// Tests for HalfBROT.FB_FocusManualHome, the decision and the end detection of a manual focus re-home, calibrated or not (HalfBROT 0.11.0, #138).
// The wiring in FB_FocusControl and the NC behaviour are not testable here (the mock skips the body): on-site test.
FUNCTION_BLOCK FB_FocusManualHome_Tests EXTENDS TcUnit.FB_TestSuite
VAR
END_VAR

Accepted_When_Calibrated_Idle_Automatic();
Rejected_In_Manual_Mode();
Rejected_With_Manual_Unlock();
Rejected_With_Axis_Error();
Accepted_When_Not_Calibrated();
Uncalibrated_Rejected_In_Manual_Mode();
Uncalibrated_Rejected_While_Homing();
Uncalibrated_Rejected_With_Error();
Uncalibrated_Rejected_With_Manual_Unlock();
Uncalibrated_Rejected_While_Moving();
NotAutomatic_Before_Homing();
No_Second_Request_While_Running_Uncalibrated();
Calibrated_Request_Restores_Target();
Uncalibrated_Done_No_Restore();
Uncalibrated_Abort_Blocks_AutoHome();
Uncalibrated_Abort_Before_Start();
Rejected_While_Homing();
Rejected_While_Moving();
No_Second_Request_While_Running();
Done_After_Active_And_Calibrated();
Done_When_Calibrated_Stays_True();
Done_When_Calibrated_Drops_And_Returns();
Abort_By_Stop_Pulse();
Abort_By_Error();
Abort_Before_Start();
Abort_Uncalibrated_Blocks_AutoHome();
Abort_Calibrated_No_Block();
Request_Clears_Block();
ClearBlock();
Aborted_Rehome_Then_Rehome_Restores_The_First_Target();
ClearBlock_Drops_The_Kept_Target();
Calibrated_Abort_Drops_The_Pending_Target();

// The plain case: accepted, running, the target is kept for the end.
METHOD PRIVATE Accepted_When_Calibrated_Idle_Automatic
VAR
	fb	: HalfBROT.FB_FocusManualHome;
	eRes	: HalfBROT.E_FocusManualHome;
END_VAR
TEST('Accepted_When_Calibrated_Idle_Automatic');
eRes := fb.Request(bAutomatic := TRUE, bManualUnlock := FALSE, bError := FALSE, bCalibrated := TRUE, bHoming := FALSE, bMoving := FALSE, fTarget := 36.0);
AssertTrue(Condition := eRes = HalfBROT.E_FocusManualHome.Accepted, Message := 'accepted');
AssertTrue(Condition := fb.bRunning, Message := 'running');
AssertFalse(Condition := fb.bBlockAutoHome, Message := 'no block');
AssertEquals_LREAL(Expected := 36.0, Actual := fb.fRestoreTarget, Delta := 1.0E-9, Message := 'target kept');
AssertTrue(Condition := fb.bRestoreTarget, Message := 'restore the target');
TEST_FINISHED();
END_METHOD

// Manual/pendant mode: the pendant drives the enable and jogs.
METHOD PRIVATE Rejected_In_Manual_Mode
VAR
	fb	: HalfBROT.FB_FocusManualHome;
	eRes	: HalfBROT.E_FocusManualHome;
END_VAR
TEST('Rejected_In_Manual_Mode');
eRes := fb.Request(bAutomatic := FALSE, bManualUnlock := FALSE, bError := FALSE, bCalibrated := TRUE, bHoming := FALSE, bMoving := FALSE, fTarget := 36.0);
AssertTrue(Condition := eRes = HalfBROT.E_FocusManualHome.NotAutomatic, Message := 'manual mode');
AssertFalse(Condition := fb.bRunning, Message := 'nothing started');
TEST_FINISHED();
END_METHOD

METHOD PRIVATE Rejected_With_Manual_Unlock
VAR
	fb	: HalfBROT.FB_FocusManualHome;
	eRes	: HalfBROT.E_FocusManualHome;
END_VAR
TEST('Rejected_With_Manual_Unlock');
eRes := fb.Request(bAutomatic := TRUE, bManualUnlock := TRUE, bError := FALSE, bCalibrated := TRUE, bHoming := FALSE, bMoving := FALSE, fTarget := 36.0);
AssertTrue(Condition := eRes = HalfBROT.E_FocusManualHome.ManualUnlock, Message := 'manual unlock');
AssertFalse(Condition := fb.bRunning, Message := 'nothing started');
TEST_FINISHED();
END_METHOD

METHOD PRIVATE Rejected_With_Axis_Error
VAR
	fb	: HalfBROT.FB_FocusManualHome;
	eRes	: HalfBROT.E_FocusManualHome;
END_VAR
TEST('Rejected_With_Axis_Error');
eRes := fb.Request(bAutomatic := TRUE, bManualUnlock := FALSE, bError := TRUE, bCalibrated := TRUE, bHoming := FALSE, bMoving := FALSE, fTarget := 36.0);
AssertTrue(Condition := eRes = HalfBROT.E_FocusManualHome.AxisError, Message := 'axis error');
AssertFalse(Condition := fb.bRunning, Message := 'nothing started');
TEST_FINISHED();
END_METHOD

// A homing is requested, pending or active (the caller passes bHomeAxis OR HomeActive OR HomePending).
METHOD PRIVATE Rejected_While_Homing
VAR
	fb	: HalfBROT.FB_FocusManualHome;
	eRes	: HalfBROT.E_FocusManualHome;
END_VAR
TEST('Rejected_While_Homing');
eRes := fb.Request(bAutomatic := TRUE, bManualUnlock := FALSE, bError := FALSE, bCalibrated := TRUE, bHoming := TRUE, bMoving := FALSE, fTarget := 36.0);
AssertTrue(Condition := eRes = HalfBROT.E_FocusManualHome.Homing, Message := 'homing');
AssertFalse(Condition := fb.bRunning, Message := 'nothing started');
TEST_FINISHED();
END_METHOD

METHOD PRIVATE Rejected_While_Moving
VAR
	fb	: HalfBROT.FB_FocusManualHome;
	eRes	: HalfBROT.E_FocusManualHome;
END_VAR
TEST('Rejected_While_Moving');
eRes := fb.Request(bAutomatic := TRUE, bManualUnlock := FALSE, bError := FALSE, bCalibrated := TRUE, bHoming := FALSE, bMoving := TRUE, fTarget := 36.0);
AssertTrue(Condition := eRes = HalfBROT.E_FocusManualHome.Moving, Message := 'moving');
AssertFalse(Condition := fb.bRunning, Message := 'nothing started');
TEST_FINISHED();
END_METHOD

METHOD PRIVATE No_Second_Request_While_Running
VAR
	fb	: HalfBROT.FB_FocusManualHome;
	eRes	: HalfBROT.E_FocusManualHome;
END_VAR
TEST('No_Second_Request_While_Running');
eRes := fb.Request(bAutomatic := TRUE, bManualUnlock := FALSE, bError := FALSE, bCalibrated := TRUE, bHoming := FALSE, bMoving := FALSE, fTarget := 36.0);
eRes := fb.Request(bAutomatic := TRUE, bManualUnlock := FALSE, bError := FALSE, bCalibrated := TRUE, bHoming := FALSE, bMoving := FALSE, fTarget := 50.0);
AssertTrue(Condition := eRes = HalfBROT.E_FocusManualHome.Homing, Message := 'second request');
AssertEquals_LREAL(Expected := 36.0, Actual := fb.fRestoreTarget, Delta := 1.0E-9, Message := 'first target kept');
TEST_FINISHED();
END_METHOD

// Pending, active, then calibrated and idle: done for one cycle, restore target available.
METHOD PRIVATE Done_After_Active_And_Calibrated
VAR
	fb	: HalfBROT.FB_FocusManualHome;
	eRes	: HalfBROT.E_FocusManualHome;
END_VAR
TEST('Done_After_Active_And_Calibrated');
eRes := fb.Request(bAutomatic := TRUE, bManualUnlock := FALSE, bError := FALSE, bCalibrated := TRUE, bHoming := FALSE, bMoving := FALSE, fTarget := 36.0);
fb(bHomeActive := FALSE, bHomePending := TRUE, bCalibrated := TRUE, bAbortPulse := FALSE);
AssertTrue(Condition := fb.bRunning, Message := 'running while pending');
fb(bHomeActive := TRUE, bHomePending := FALSE, bCalibrated := TRUE, bAbortPulse := FALSE);
AssertTrue(Condition := fb.bRunning, Message := 'running while active');
AssertFalse(Condition := fb.bDone, Message := 'not done yet');
fb(bHomeActive := FALSE, bHomePending := FALSE, bCalibrated := TRUE, bAbortPulse := FALSE);
AssertTrue(Condition := fb.bDone, Message := 'done');
AssertFalse(Condition := fb.bRunning, Message := 'ended');
AssertFalse(Condition := fb.bAborted, Message := 'not aborted');
AssertFalse(Condition := fb.bBlockAutoHome, Message := 'no block');
fb(bHomeActive := FALSE, bHomePending := FALSE, bCalibrated := TRUE, bAbortPulse := FALSE);
AssertFalse(Condition := fb.bDone, Message := 'done is one cycle');
TEST_FINISHED();
END_METHOD

// The NC keeps Homed during the homing.
METHOD PRIVATE Done_When_Calibrated_Stays_True
VAR
	fb	: HalfBROT.FB_FocusManualHome;
	eRes	: HalfBROT.E_FocusManualHome;
END_VAR
TEST('Done_When_Calibrated_Stays_True');
eRes := fb.Request(bAutomatic := TRUE, bManualUnlock := FALSE, bError := FALSE, bCalibrated := TRUE, bHoming := FALSE, bMoving := FALSE, fTarget := 36.0);
fb(bHomeActive := TRUE, bHomePending := FALSE, bCalibrated := TRUE, bAbortPulse := FALSE);
fb(bHomeActive := TRUE, bHomePending := FALSE, bCalibrated := TRUE, bAbortPulse := FALSE);
fb(bHomeActive := FALSE, bHomePending := FALSE, bCalibrated := TRUE, bAbortPulse := FALSE);
AssertTrue(Condition := fb.bDone, Message := 'done');
TEST_FINISHED();
END_METHOD

// The NC drops Homed at the start of the homing.
METHOD PRIVATE Done_When_Calibrated_Drops_And_Returns
VAR
	fb	: HalfBROT.FB_FocusManualHome;
	eRes	: HalfBROT.E_FocusManualHome;
END_VAR
TEST('Done_When_Calibrated_Drops_And_Returns');
eRes := fb.Request(bAutomatic := TRUE, bManualUnlock := FALSE, bError := FALSE, bCalibrated := TRUE, bHoming := FALSE, bMoving := FALSE, fTarget := 36.0);
fb(bHomeActive := FALSE, bHomePending := TRUE, bCalibrated := TRUE, bAbortPulse := FALSE);
fb(bHomeActive := TRUE, bHomePending := FALSE, bCalibrated := FALSE, bAbortPulse := FALSE);
fb(bHomeActive := TRUE, bHomePending := FALSE, bCalibrated := FALSE, bAbortPulse := FALSE);
fb(bHomeActive := FALSE, bHomePending := FALSE, bCalibrated := TRUE, bAbortPulse := FALSE);
AssertTrue(Condition := fb.bDone, Message := 'done');
AssertFalse(Condition := fb.bBlockAutoHome, Message := 'no block');
TEST_FINISHED();
END_METHOD

// A stop aborts the homing; the axis keeps its old calibration.
METHOD PRIVATE Abort_By_Stop_Pulse
VAR
	fb	: HalfBROT.FB_FocusManualHome;
	eRes	: HalfBROT.E_FocusManualHome;
END_VAR
TEST('Abort_By_Stop_Pulse');
eRes := fb.Request(bAutomatic := TRUE, bManualUnlock := FALSE, bError := FALSE, bCalibrated := TRUE, bHoming := FALSE, bMoving := FALSE, fTarget := 36.0);
fb(bHomeActive := TRUE, bHomePending := FALSE, bCalibrated := TRUE, bAbortPulse := FALSE);
fb(bHomeActive := TRUE, bHomePending := FALSE, bCalibrated := TRUE, bAbortPulse := TRUE);
fb(bHomeActive := FALSE, bHomePending := FALSE, bCalibrated := TRUE, bAbortPulse := FALSE);
AssertTrue(Condition := fb.bAborted, Message := 'aborted');
AssertFalse(Condition := fb.bDone, Message := 'not done');
AssertFalse(Condition := fb.bRunning, Message := 'ended');
AssertFalse(Condition := fb.bBlockAutoHome, Message := 'calibrated: no block');
TEST_FINISHED();
END_METHOD

// An axis error ends the homing uncalibrated.
METHOD PRIVATE Abort_By_Error
VAR
	fb	: HalfBROT.FB_FocusManualHome;
	eRes	: HalfBROT.E_FocusManualHome;
END_VAR
TEST('Abort_By_Error');
eRes := fb.Request(bAutomatic := TRUE, bManualUnlock := FALSE, bError := FALSE, bCalibrated := TRUE, bHoming := FALSE, bMoving := FALSE, fTarget := 36.0);
fb(bHomeActive := TRUE, bHomePending := FALSE, bCalibrated := TRUE, bAbortPulse := FALSE);
fb(bHomeActive := TRUE, bHomePending := FALSE, bCalibrated := FALSE, bAbortPulse := TRUE);
fb(bHomeActive := FALSE, bHomePending := FALSE, bCalibrated := FALSE, bAbortPulse := FALSE);
AssertTrue(Condition := fb.bAborted, Message := 'aborted');
AssertFalse(Condition := fb.bDone, Message := 'not done');
AssertTrue(Condition := fb.bBlockAutoHome, Message := 'uncalibrated: block');
TEST_FINISHED();
END_METHOD

// Stop() cancels a Home() that still waits for the drive: HomeActive is never seen.
METHOD PRIVATE Abort_Before_Start
VAR
	fb	: HalfBROT.FB_FocusManualHome;
	eRes	: HalfBROT.E_FocusManualHome;
END_VAR
TEST('Abort_Before_Start');
eRes := fb.Request(bAutomatic := TRUE, bManualUnlock := FALSE, bError := FALSE, bCalibrated := TRUE, bHoming := FALSE, bMoving := FALSE, fTarget := 36.0);
fb(bHomeActive := FALSE, bHomePending := TRUE, bCalibrated := TRUE, bAbortPulse := FALSE);
fb(bHomeActive := FALSE, bHomePending := FALSE, bCalibrated := TRUE, bAbortPulse := FALSE);
AssertTrue(Condition := fb.bAborted, Message := 'aborted');
AssertFalse(Condition := fb.bDone, Message := 'not done: never active');
AssertFalse(Condition := fb.bBlockAutoHome, Message := 'calibrated: no block');
TEST_FINISHED();
END_METHOD

// Ends uncalibrated: the automatic homing stays off.
METHOD PRIVATE Abort_Uncalibrated_Blocks_AutoHome
VAR
	fb	: HalfBROT.FB_FocusManualHome;
	eRes	: HalfBROT.E_FocusManualHome;
END_VAR
TEST('Abort_Uncalibrated_Blocks_AutoHome');
eRes := fb.Request(bAutomatic := TRUE, bManualUnlock := FALSE, bError := FALSE, bCalibrated := TRUE, bHoming := FALSE, bMoving := FALSE, fTarget := 36.0);
fb(bHomeActive := TRUE, bHomePending := FALSE, bCalibrated := FALSE, bAbortPulse := FALSE);
fb(bHomeActive := FALSE, bHomePending := FALSE, bCalibrated := FALSE, bAbortPulse := FALSE);
AssertTrue(Condition := fb.bAborted, Message := 'aborted');
AssertTrue(Condition := fb.bBlockAutoHome, Message := 'block');
TEST_FINISHED();
END_METHOD

METHOD PRIVATE Abort_Calibrated_No_Block
VAR
	fb	: HalfBROT.FB_FocusManualHome;
	eRes	: HalfBROT.E_FocusManualHome;
END_VAR
TEST('Abort_Calibrated_No_Block');
eRes := fb.Request(bAutomatic := TRUE, bManualUnlock := FALSE, bError := FALSE, bCalibrated := TRUE, bHoming := FALSE, bMoving := FALSE, fTarget := 36.0);
fb(bHomeActive := TRUE, bHomePending := FALSE, bCalibrated := TRUE, bAbortPulse := FALSE);
fb(bHomeActive := TRUE, bHomePending := FALSE, bCalibrated := TRUE, bAbortPulse := TRUE);
fb(bHomeActive := FALSE, bHomePending := FALSE, bCalibrated := TRUE, bAbortPulse := FALSE);
AssertFalse(Condition := fb.bBlockAutoHome, Message := 'no block');
TEST_FINISHED();
END_METHOD

// An uncalibrated focus is accepted while the automatic homing is blocked, and the request lifts the block.
// The target of the aborted re-home before it is kept (HalfBROT#152; was: no target to restore).
METHOD PRIVATE Request_Clears_Block
VAR
	fb	: HalfBROT.FB_FocusManualHome;
	eRes	: HalfBROT.E_FocusManualHome;
END_VAR
TEST('Request_Clears_Block');
eRes := fb.Request(bAutomatic := TRUE, bManualUnlock := FALSE, bError := FALSE, bCalibrated := TRUE, bHoming := FALSE, bMoving := FALSE, fTarget := 36.0);
fb(bHomeActive := TRUE, bHomePending := FALSE, bCalibrated := FALSE, bAbortPulse := FALSE);
fb(bHomeActive := FALSE, bHomePending := FALSE, bCalibrated := FALSE, bAbortPulse := FALSE);
eRes := fb.Request(bAutomatic := TRUE, bManualUnlock := FALSE, bError := FALSE, bCalibrated := FALSE, bHoming := FALSE, bMoving := FALSE, fTarget := 36.0);
AssertTrue(Condition := eRes = HalfBROT.E_FocusManualHome.Accepted, Message := 'accepted while blocked');
AssertFalse(Condition := fb.bBlockAutoHome, Message := 'block lifted');
AssertTrue(Condition := fb.bRunning, Message := 'running');
AssertTrue(Condition := fb.bRestoreTarget, Message := 'the target of the aborted re-home is kept (#152)');
AssertEquals_LREAL(Expected := 36.0, Actual := fb.fRestoreTarget, Delta := 1.0E-9, Message := 'first target, not the junk one');
TEST_FINISHED();
END_METHOD

// Another homing request lifts the block.
METHOD PRIVATE ClearBlock
VAR
	fb	: HalfBROT.FB_FocusManualHome;
	eRes	: HalfBROT.E_FocusManualHome;
END_VAR
TEST('ClearBlock');
eRes := fb.Request(bAutomatic := TRUE, bManualUnlock := FALSE, bError := FALSE, bCalibrated := TRUE, bHoming := FALSE, bMoving := FALSE, fTarget := 36.0);
fb(bHomeActive := TRUE, bHomePending := FALSE, bCalibrated := FALSE, bAbortPulse := FALSE);
fb(bHomeActive := FALSE, bHomePending := FALSE, bCalibrated := FALSE, bAbortPulse := FALSE);
AssertTrue(Condition := fb.bBlockAutoHome, Message := 'block');
fb.ClearBlock();
AssertFalse(Condition := fb.bBlockAutoHome, Message := 'cleared');
TEST_FINISHED();
END_METHOD

// HalfBROT#152 (MS-135): a stop in the sweep of a re-home from 35.98 mm, then bManualHome again to the end.
// The second request is on an uncalibrated focus (fTarget is junk there, 0 in MS-135) and must still restore 35.98.
// The target is used up by the cycle of bDone; a later request on the uncalibrated focus has none.
METHOD PRIVATE Aborted_Rehome_Then_Rehome_Restores_The_First_Target
VAR
	fb	: HalfBROT.FB_FocusManualHome;
	eRes	: HalfBROT.E_FocusManualHome;
END_VAR
TEST('Aborted_Rehome_Then_Rehome_Restores_The_First_Target');
eRes := fb.Request(bAutomatic := TRUE, bManualUnlock := FALSE, bError := FALSE, bCalibrated := TRUE, bHoming := FALSE, bMoving := FALSE, fTarget := 35.98);
fb(bHomeActive := TRUE, bHomePending := FALSE, bCalibrated := FALSE, bAbortPulse := FALSE);
fb(bHomeActive := TRUE, bHomePending := FALSE, bCalibrated := FALSE, bAbortPulse := TRUE);
fb(bHomeActive := FALSE, bHomePending := FALSE, bCalibrated := FALSE, bAbortPulse := FALSE);
AssertTrue(Condition := fb.bAborted, Message := 'first re-home aborted');
AssertTrue(Condition := fb.bBlockAutoHome, Message := 'blocked, uncalibrated');
eRes := fb.Request(bAutomatic := TRUE, bManualUnlock := FALSE, bError := FALSE, bCalibrated := FALSE, bHoming := FALSE, bMoving := FALSE, fTarget := 0.0);
AssertTrue(Condition := eRes = HalfBROT.E_FocusManualHome.Accepted, Message := 'second accepted');
AssertTrue(Condition := fb.bRestoreTarget, Message := 'restore pending');
AssertEquals_LREAL(Expected := 35.98, Actual := fb.fRestoreTarget, Delta := 1.0E-9, Message := 'first target kept');
fb(bHomeActive := FALSE, bHomePending := TRUE, bCalibrated := FALSE, bAbortPulse := FALSE);
fb(bHomeActive := TRUE, bHomePending := FALSE, bCalibrated := FALSE, bAbortPulse := FALSE);
fb(bHomeActive := TRUE, bHomePending := FALSE, bCalibrated := TRUE, bAbortPulse := FALSE);
fb(bHomeActive := FALSE, bHomePending := FALSE, bCalibrated := TRUE, bAbortPulse := FALSE);
AssertTrue(Condition := fb.bDone, Message := 'second re-home done');
AssertTrue(Condition := fb.bRestoreTarget, Message := 'target still there in the cycle of bDone');
AssertEquals_LREAL(Expected := 35.98, Actual := fb.fRestoreTarget, Delta := 1.0E-9, Message := 'restore 35.98');
fb(bHomeActive := FALSE, bHomePending := FALSE, bCalibrated := TRUE, bAbortPulse := FALSE);
AssertFalse(Condition := fb.bRestoreTarget, Message := 'used up the cycle after');
eRes := fb.Request(bAutomatic := TRUE, bManualUnlock := FALSE, bError := FALSE, bCalibrated := FALSE, bHoming := FALSE, bMoving := FALSE, fTarget := 12.0);
AssertFalse(Condition := fb.bRestoreTarget, Message := 'a later uncalibrated request has none');
TEST_FINISHED();
END_METHOD

// Another homing request (the power-on homing) lifts the block and ends on the cam without a restore:
// a target kept from an aborted re-home is stale then (HalfBROT#152).
METHOD PRIVATE ClearBlock_Drops_The_Kept_Target
VAR
	fb	: HalfBROT.FB_FocusManualHome;
	eRes	: HalfBROT.E_FocusManualHome;
END_VAR
TEST('ClearBlock_Drops_The_Kept_Target');
eRes := fb.Request(bAutomatic := TRUE, bManualUnlock := FALSE, bError := FALSE, bCalibrated := TRUE, bHoming := FALSE, bMoving := FALSE, fTarget := 35.98);
fb(bHomeActive := TRUE, bHomePending := FALSE, bCalibrated := FALSE, bAbortPulse := FALSE);
fb(bHomeActive := FALSE, bHomePending := FALSE, bCalibrated := FALSE, bAbortPulse := FALSE);
AssertTrue(Condition := fb.bBlockAutoHome, Message := 'blocked');
fb.ClearBlock();
eRes := fb.Request(bAutomatic := TRUE, bManualUnlock := FALSE, bError := FALSE, bCalibrated := FALSE, bHoming := FALSE, bMoving := FALSE, fTarget := 0.0);
AssertTrue(Condition := eRes = HalfBROT.E_FocusManualHome.Accepted, Message := 'accepted');
AssertFalse(Condition := fb.bRestoreTarget, Message := 'no stale target');
AssertEquals_LREAL(Expected := 0.0, Actual := fb.fRestoreTarget, Delta := 1.0E-9, Message := 'no junk target kept');
TEST_FINISHED();
END_METHOD

// A stop that leaves the calibration alone ends the re-home for good: nothing stays pending for a later uncalibrated request.
METHOD PRIVATE Calibrated_Abort_Drops_The_Pending_Target
VAR
	fb	: HalfBROT.FB_FocusManualHome;
	eRes	: HalfBROT.E_FocusManualHome;
END_VAR
TEST('Calibrated_Abort_Drops_The_Pending_Target');
eRes := fb.Request(bAutomatic := TRUE, bManualUnlock := FALSE, bError := FALSE, bCalibrated := TRUE, bHoming := FALSE, bMoving := FALSE, fTarget := 35.98);
fb(bHomeActive := TRUE, bHomePending := FALSE, bCalibrated := TRUE, bAbortPulse := FALSE);
fb(bHomeActive := TRUE, bHomePending := FALSE, bCalibrated := TRUE, bAbortPulse := TRUE);
fb(bHomeActive := FALSE, bHomePending := FALSE, bCalibrated := TRUE, bAbortPulse := FALSE);
AssertTrue(Condition := fb.bAborted, Message := 'aborted');
AssertFalse(Condition := fb.bBlockAutoHome, Message := 'calibrated: no block');
AssertFalse(Condition := fb.bRestoreTarget, Message := 'nothing pending');
eRes := fb.Request(bAutomatic := TRUE, bManualUnlock := FALSE, bError := FALSE, bCalibrated := FALSE, bHoming := FALSE, bMoving := FALSE, fTarget := 12.0);
AssertFalse(Condition := fb.bRestoreTarget, Message := 'a later uncalibrated request has none');
TEST_FINISHED();
END_METHOD

// An uncalibrated focus is accepted (#138): no target to restore, fPosition is junk there (#115).
METHOD PRIVATE Accepted_When_Not_Calibrated
VAR
	fb	: HalfBROT.FB_FocusManualHome;
	eRes	: HalfBROT.E_FocusManualHome;
END_VAR
TEST('Accepted_When_Not_Calibrated');
eRes := fb.Request(bAutomatic := TRUE, bManualUnlock := FALSE, bError := FALSE, bCalibrated := FALSE, bHoming := FALSE, bMoving := FALSE, fTarget := 36.0);
AssertTrue(Condition := eRes = HalfBROT.E_FocusManualHome.Accepted, Message := 'accepted');
AssertTrue(Condition := fb.bRunning, Message := 'running');
AssertFalse(Condition := fb.bRestoreTarget, Message := 'no target to restore');
AssertFalse(Condition := fb.bBlockAutoHome, Message := 'no block');
TEST_FINISHED();
END_METHOD

// Manual mode stays refused: the drive is only enabled in automatic.
METHOD PRIVATE Uncalibrated_Rejected_In_Manual_Mode
VAR
	fb	: HalfBROT.FB_FocusManualHome;
	eRes	: HalfBROT.E_FocusManualHome;
END_VAR
TEST('Uncalibrated_Rejected_In_Manual_Mode');
eRes := fb.Request(bAutomatic := FALSE, bManualUnlock := FALSE, bError := FALSE, bCalibrated := FALSE, bHoming := FALSE, bMoving := FALSE, fTarget := 36.0);
AssertTrue(Condition := eRes = HalfBROT.E_FocusManualHome.NotAutomatic, Message := 'manual mode');
AssertFalse(Condition := fb.bRunning, Message := 'nothing started');
TEST_FINISHED();
END_METHOD

// The automatic homing was already requested: the request is refused.
METHOD PRIVATE Uncalibrated_Rejected_While_Homing
VAR
	fb	: HalfBROT.FB_FocusManualHome;
	eRes	: HalfBROT.E_FocusManualHome;
END_VAR
TEST('Uncalibrated_Rejected_While_Homing');
eRes := fb.Request(bAutomatic := TRUE, bManualUnlock := FALSE, bError := FALSE, bCalibrated := FALSE, bHoming := TRUE, bMoving := FALSE, fTarget := 36.0);
AssertTrue(Condition := eRes = HalfBROT.E_FocusManualHome.Homing, Message := 'homing');
AssertFalse(Condition := fb.bRunning, Message := 'nothing started');
TEST_FINISHED();
END_METHOD

// The checks before the acceptance still apply.
METHOD PRIVATE Uncalibrated_Rejected_With_Error
VAR
	fb	: HalfBROT.FB_FocusManualHome;
	eRes	: HalfBROT.E_FocusManualHome;
END_VAR
TEST('Uncalibrated_Rejected_With_Error');
eRes := fb.Request(bAutomatic := TRUE, bManualUnlock := FALSE, bError := TRUE, bCalibrated := FALSE, bHoming := FALSE, bMoving := FALSE, fTarget := 36.0);
AssertTrue(Condition := eRes = HalfBROT.E_FocusManualHome.AxisError, Message := 'axis error');
AssertFalse(Condition := fb.bRunning, Message := 'nothing started');
TEST_FINISHED();
END_METHOD

// The checks before the acceptance still apply.
METHOD PRIVATE Uncalibrated_Rejected_With_Manual_Unlock
VAR
	fb	: HalfBROT.FB_FocusManualHome;
	eRes	: HalfBROT.E_FocusManualHome;
END_VAR
TEST('Uncalibrated_Rejected_With_Manual_Unlock');
eRes := fb.Request(bAutomatic := TRUE, bManualUnlock := TRUE, bError := FALSE, bCalibrated := FALSE, bHoming := FALSE, bMoving := FALSE, fTarget := 36.0);
AssertTrue(Condition := eRes = HalfBROT.E_FocusManualHome.ManualUnlock, Message := 'manual unlock');
AssertFalse(Condition := fb.bRunning, Message := 'nothing started');
TEST_FINISHED();
END_METHOD

// The checks before the acceptance still apply.
METHOD PRIVATE Uncalibrated_Rejected_While_Moving
VAR
	fb	: HalfBROT.FB_FocusManualHome;
	eRes	: HalfBROT.E_FocusManualHome;
END_VAR
TEST('Uncalibrated_Rejected_While_Moving');
eRes := fb.Request(bAutomatic := TRUE, bManualUnlock := FALSE, bError := FALSE, bCalibrated := FALSE, bHoming := FALSE, bMoving := TRUE, fTarget := 36.0);
AssertTrue(Condition := eRes = HalfBROT.E_FocusManualHome.Moving, Message := 'moving');
AssertFalse(Condition := fb.bRunning, Message := 'nothing started');
TEST_FINISHED();
END_METHOD

// Priority: manual mode is reported before a running homing.
METHOD PRIVATE NotAutomatic_Before_Homing
VAR
	fb	: HalfBROT.FB_FocusManualHome;
	eRes	: HalfBROT.E_FocusManualHome;
END_VAR
TEST('NotAutomatic_Before_Homing');
eRes := fb.Request(bAutomatic := FALSE, bManualUnlock := FALSE, bError := FALSE, bCalibrated := FALSE, bHoming := TRUE, bMoving := FALSE, fTarget := 36.0);
AssertTrue(Condition := eRes = HalfBROT.E_FocusManualHome.NotAutomatic, Message := 'manual mode first');
TEST_FINISHED();
END_METHOD

// A doubled Start is refused and the first request is kept.
METHOD PRIVATE No_Second_Request_While_Running_Uncalibrated
VAR
	fb	: HalfBROT.FB_FocusManualHome;
	eRes	: HalfBROT.E_FocusManualHome;
END_VAR
TEST('No_Second_Request_While_Running_Uncalibrated');
eRes := fb.Request(bAutomatic := TRUE, bManualUnlock := FALSE, bError := FALSE, bCalibrated := FALSE, bHoming := FALSE, bMoving := FALSE, fTarget := 36.0);
eRes := fb.Request(bAutomatic := TRUE, bManualUnlock := FALSE, bError := FALSE, bCalibrated := FALSE, bHoming := FALSE, bMoving := FALSE, fTarget := 50.0);
AssertTrue(Condition := eRes = HalfBROT.E_FocusManualHome.Homing, Message := 'second request');
AssertFalse(Condition := fb.bRestoreTarget, Message := 'still no target');
AssertEquals_LREAL(Expected := 0.0, Actual := fb.fRestoreTarget, Delta := 1.0E-9, Message := 'no junk target kept');
TEST_FINISHED();
END_METHOD

// A request on a calibrated focus keeps its target for the end.
METHOD PRIVATE Calibrated_Request_Restores_Target
VAR
	fb	: HalfBROT.FB_FocusManualHome;
	eRes	: HalfBROT.E_FocusManualHome;
END_VAR
TEST('Calibrated_Request_Restores_Target');
eRes := fb.Request(bAutomatic := TRUE, bManualUnlock := FALSE, bError := FALSE, bCalibrated := TRUE, bHoming := FALSE, bMoving := FALSE, fTarget := 36.0);
AssertTrue(Condition := fb.bRestoreTarget, Message := 'restore the target');
AssertEquals_LREAL(Expected := 36.0, Actual := fb.fRestoreTarget, Delta := 1.0E-9, Message := 'target kept');
TEST_FINISHED();
END_METHOD

// Pending, active, then calibrated and idle: done, nothing to restore.
METHOD PRIVATE Uncalibrated_Done_No_Restore
VAR
	fb	: HalfBROT.FB_FocusManualHome;
	eRes	: HalfBROT.E_FocusManualHome;
END_VAR
TEST('Uncalibrated_Done_No_Restore');
eRes := fb.Request(bAutomatic := TRUE, bManualUnlock := FALSE, bError := FALSE, bCalibrated := FALSE, bHoming := FALSE, bMoving := FALSE, fTarget := 36.0);
fb(bHomeActive := FALSE, bHomePending := TRUE, bCalibrated := FALSE, bAbortPulse := FALSE);
fb(bHomeActive := TRUE, bHomePending := FALSE, bCalibrated := FALSE, bAbortPulse := FALSE);
fb(bHomeActive := TRUE, bHomePending := FALSE, bCalibrated := TRUE, bAbortPulse := FALSE);
fb(bHomeActive := FALSE, bHomePending := FALSE, bCalibrated := TRUE, bAbortPulse := FALSE);
AssertTrue(Condition := fb.bDone, Message := 'done');
AssertFalse(Condition := fb.bAborted, Message := 'not aborted');
AssertFalse(Condition := fb.bBlockAutoHome, Message := 'no block');
AssertFalse(Condition := fb.bRestoreTarget, Message := 'no restore');
TEST_FINISHED();
END_METHOD

// A stop during an uncalibrated homing: aborted, the automatic homing stays off.
METHOD PRIVATE Uncalibrated_Abort_Blocks_AutoHome
VAR
	fb	: HalfBROT.FB_FocusManualHome;
	eRes	: HalfBROT.E_FocusManualHome;
END_VAR
TEST('Uncalibrated_Abort_Blocks_AutoHome');
eRes := fb.Request(bAutomatic := TRUE, bManualUnlock := FALSE, bError := FALSE, bCalibrated := FALSE, bHoming := FALSE, bMoving := FALSE, fTarget := 36.0);
fb(bHomeActive := TRUE, bHomePending := FALSE, bCalibrated := FALSE, bAbortPulse := FALSE);
fb(bHomeActive := TRUE, bHomePending := FALSE, bCalibrated := FALSE, bAbortPulse := TRUE);
fb(bHomeActive := FALSE, bHomePending := FALSE, bCalibrated := FALSE, bAbortPulse := FALSE);
AssertTrue(Condition := fb.bAborted, Message := 'aborted');
AssertFalse(Condition := fb.bDone, Message := 'not done');
AssertTrue(Condition := fb.bBlockAutoHome, Message := 'block');
TEST_FINISHED();
END_METHOD

// Stop() cancels a Home() that waits for the drive: never active, aborted, blocked.
METHOD PRIVATE Uncalibrated_Abort_Before_Start
VAR
	fb	: HalfBROT.FB_FocusManualHome;
	eRes	: HalfBROT.E_FocusManualHome;
END_VAR
TEST('Uncalibrated_Abort_Before_Start');
eRes := fb.Request(bAutomatic := TRUE, bManualUnlock := FALSE, bError := FALSE, bCalibrated := FALSE, bHoming := FALSE, bMoving := FALSE, fTarget := 36.0);
fb(bHomeActive := FALSE, bHomePending := TRUE, bCalibrated := FALSE, bAbortPulse := FALSE);
fb(bHomeActive := FALSE, bHomePending := FALSE, bCalibrated := FALSE, bAbortPulse := FALSE);
AssertTrue(Condition := fb.bAborted, Message := 'aborted');
AssertFalse(Condition := fb.bDone, Message := 'not done: never active');
AssertTrue(Condition := fb.bBlockAutoHome, Message := 'block');
TEST_FINISHED();
END_METHOD

END_FUNCTION_BLOCK

(* stored: Version 1.1.0.1, ProductVersion 3.1.4024.15
   POU FB_FocusManualHome_Tests: Id {0817fa45-2195-4f20-91e2-fdb09ceb798d}, SpecialFunc None
   Method Accepted_When_Calibrated_Idle_Automatic: Id {1ff9da75-f12f-4899-bc74-50b4fb651ac8}
   Method Rejected_In_Manual_Mode: Id {e4aa7f98-bc8e-4d12-8ae5-d32033812655}
   Method Rejected_With_Manual_Unlock: Id {e9a3b0e6-9532-4423-9f0b-0f8b6d1b2110}
   Method Rejected_With_Axis_Error: Id {6f8609dd-6f06-405a-ae1b-b36b5911a5b7}
   Method Rejected_While_Homing: Id {9eb6bd9d-0758-48b3-88fc-f185ded4ec4b}
   Method Rejected_While_Moving: Id {152bef88-baa1-4048-93ef-4014528f23d1}
   Method No_Second_Request_While_Running: Id {08c47c24-3cdf-44a1-af1e-31667849e213}
   Method Done_After_Active_And_Calibrated: Id {0ef3ac99-9e51-4436-9c3d-9254f85fca07}
   Method Done_When_Calibrated_Stays_True: Id {eecd2123-600d-4994-947c-b670921f7d43}
   Method Done_When_Calibrated_Drops_And_Returns: Id {9bf78ece-46e9-4478-a30e-ff1daf0fad1b}
   Method Abort_By_Stop_Pulse: Id {e5e286bb-6208-4c6a-ba08-e2517641cefb}
   Method Abort_By_Error: Id {3e599098-3f13-45f8-b159-4e63a5c9d89b}
   Method Abort_Before_Start: Id {26270119-cce3-42d4-aa19-7ca8dfd6b8e3}
   Method Abort_Uncalibrated_Blocks_AutoHome: Id {1f3bf5f4-ac64-409a-b9d9-a6094de475d1}
   Method Abort_Calibrated_No_Block: Id {02a0766d-2a5d-4329-bd43-9efc37ddf683}
   Method Request_Clears_Block: Id {11b585a2-05af-45ef-b08d-f700249ddb87}
   Method ClearBlock: Id {42a5b9f7-e78d-40e2-9590-75912cdd3f76}
   Method Aborted_Rehome_Then_Rehome_Restores_The_First_Target: Id {3c8d1f52-7a40-4b19-9e63-0d52a7c4e8b1}
   Method ClearBlock_Drops_The_Kept_Target: Id {b7e24a90-1d6c-4f83-a5b2-9c0e3f71d6a4}
   Method Calibrated_Abort_Drops_The_Pending_Target: Id {d41a6e08-52f7-4c3b-8e19-6a0b9d2c7f35}
   Method Accepted_When_Not_Calibrated: Id {a3001c94-58ca-4dce-9d09-f28ec50baad7}
   Method Uncalibrated_Rejected_In_Manual_Mode: Id {79806093-271d-4703-8a65-023d75ab3d02}
   Method Uncalibrated_Rejected_While_Homing: Id {a06b993f-dc3c-4532-8059-c0023594597b}
   Method Uncalibrated_Rejected_With_Error: Id {2f9f5488-d7b3-48aa-a0c6-4d100b99d905}
   Method Uncalibrated_Rejected_With_Manual_Unlock: Id {7aa45950-6016-4606-ac65-e878cef48129}
   Method Uncalibrated_Rejected_While_Moving: Id {a1241849-47bf-4806-a215-3a564b8fdb8c}
   Method NotAutomatic_Before_Homing: Id {fbbc905a-8a7b-4bae-81d0-797435a25854}
   Method No_Second_Request_While_Running_Uncalibrated: Id {941d1345-f033-4b9b-a803-152d47a402cc}
   Method Calibrated_Request_Restores_Target: Id {346d1933-320b-4f57-81fd-21fb0d003118}
   Method Uncalibrated_Done_No_Restore: Id {6296907d-41bf-4dc3-9728-18dea77f3b27}
   Method Uncalibrated_Abort_Blocks_AutoHome: Id {1fbb80e5-38c9-4f7c-a6e2-bb46173ad65b}
   Method Uncalibrated_Abort_Before_Start: Id {b01c3621-de5c-4a89-89f5-b0495d65e4c1} *)
